FUNCTION_BLOCK FB_Location_Workshop
VAR_INPUT
    stInputs : ST_WorkshopInputs;
    stCommand : ST_LightCommand;
END_VAR

VAR_OUTPUT
    stOutputs : ST_WorkshopOutputs;
    stLight : ST_LightInfo;
END_VAR

VAR CONSTANT
    cLocationId : STRING(16) := 'H.01-09';
    {attribute 'TcEncoding' := 'UTF-8'}
    cLocationName : STRING(64) := UTF8#'Warsztat';
    cMainLightId : STRING(16) := 'main';
    {attribute 'TcEncoding' := 'UTF-8'}
    cMainLightName : STRING(64) := UTF8#'Oświetlenie główne';
END_VAR

VAR
    fbWorkshop : FB_ButtonLight;
END_VAR

fbWorkshop(
    bButton := stInputs.bButton,
    bAdditionalButton := FALSE,
    bSetValid := stCommand.bValid AND (stCommand.sLocationId = cLocationId) AND (stCommand.sLightId = cMainLightId),
    bTargetOn := stCommand.bTargetOn,
    bLightRelay => stOutputs.bLightRelay
);

stLight.sLocationId := cLocationId;
stLight.sLocationName := cLocationName;
stLight.sId := cMainLightId;
stLight.sName := cMainLightName;
stLight.bOn := stOutputs.bLightRelay;

END_FUNCTION_BLOCK

(* stored: Version 1.1.0.1
   POU FB_Location_Workshop: Id {ed6140a9-7ba0-4913-8278-e47fbcd68c6d}, SpecialFunc None *)
